FUNCTION_BLOCK LINEAR_START
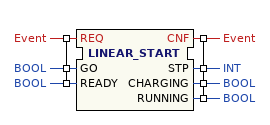
  EVENT_INPUT
    REQ WITH GO, READY;
  END_EVENT
  EVENT_OUTPUT
    CNF WITH STP, CHARGING, RUNNING;
  END_EVENT
  VAR_INPUT
    GO : BOOL;
    READY : BOOL;
  END_VAR
  VAR_OUTPUT
    STP : INT;
    CHARGING : BOOL;
    RUNNING : BOOL;
  END_VAR
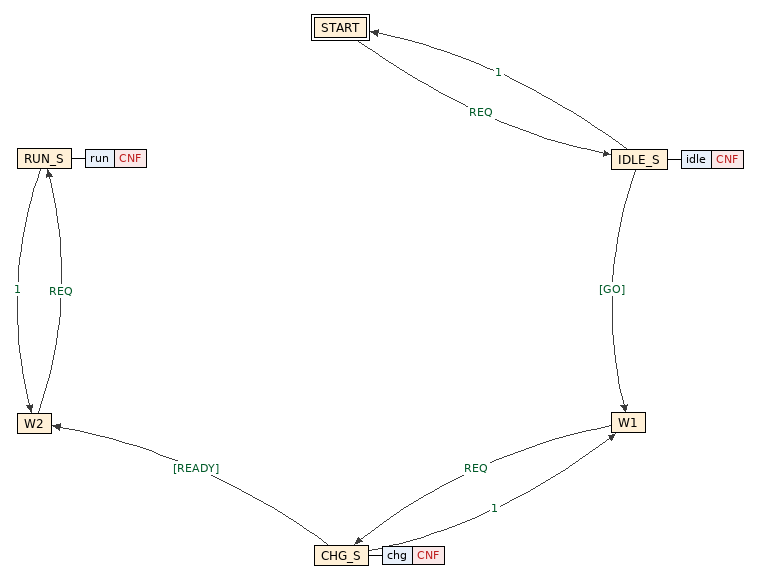
  EC_STATES
    START;
    IDLE_S : idle -> CNF;
    W1;
    CHG_S : chg -> CNF;
    W2;
    RUN_S : run -> CNF;
  END_STATES
  EC_TRANSITIONS
    START TO IDLE_S := REQ;
    IDLE_S TO W1 := [GO];
    IDLE_S TO START := 1;
    W1 TO CHG_S := REQ;
    CHG_S TO W2 := [READY];
    CHG_S TO W1 := 1;
    W2 TO RUN_S := REQ;
    RUN_S TO W2 := 1;
  END_TRANSITIONS
  ALGORITHM idle IN ST:
CHARGING := FALSE;
IF GO THEN STP := 1; END_IF;
  END_ALGORITHM
  ALGORITHM chg IN ST:
CHARGING := TRUE;
IF READY THEN STP := 2; END_IF;
  END_ALGORITHM
  ALGORITHM run IN ST:
CHARGING := FALSE;
RUNNING := TRUE;
  END_ALGORITHM
END_FUNCTION_BLOCK
